Fanuc KAREL source: KB00051.KL

PROGRAM KB00051
%NOLOCKGROUP
VAR
  P1: INTEGER
  P2: INTEGER
  RESULT: JOINTPOS
BEGIN
  P1 = 1
  P2 = 1
  RESULT = CURJPOS(P1, P2)
END KB00051
